PROGRAM MAIN
VAR
	example : FB_Example;
	filler : ARRAY[0..130] OF FB_Example;
	
	wroteData : BOOL;
	loadedData : BOOL;
END_VAR
VAR PERSISTENT
	per_example : FB_Example;
END_VAR

END_PROGRAM

(* stored: Version 1.1.0.1
   POU MAIN: Id {9cbcfa1e-4c83-4412-9b51-508f27990c15}, SpecialFunc None *)
